(*
SPDX-FileCopyrightText: c 2026 Oleksandr Tiutyk <trofimich@gmail.com>
SPDX-License-Identifier: MIT
License: https://opensource.org/license/mit
*)

(*!
<summary>Groups fixed-capacity list copying, borrowing, editing, search, sorting and overflow cases.</summary>
<description>
Owns the cases, their fixed registration array and any fixtures borrowed by the cases.
Each borrowed fixture is reserved for its case throughout the group lifetime. Use from one task at a stable address.
</description>
*)

{attribute 'no_assign'}
{attribute 'no_explicit_call' := 'do not call this function block directly'}
FUNCTION_BLOCK StaticListTestGroup EXTENDS TOF_Testing.TestGroup<16>
VAR_STAT
	{attribute 'hide'}
	_ClassName : STRING := __POUNAME();
END_VAR
VAR
	_AppendList : TOF_Collections.List<8>(valueValidator := 0);
	_InsertList : TOF_Collections.List<8>(valueValidator := 0);
	_GetAndSetList : TOF_Collections.List<8>(valueValidator := 0);
	_FindList : TOF_Collections.List<8>(valueValidator := 0);
	_ContainsList : TOF_Collections.List<8>(valueValidator := 0);
	_ContainsGenericList : TOF_Collections.List<8>(valueValidator := 0);
	_RemoveFirstList : TOF_Collections.List<8>(valueValidator := 0);
	_RemoveMatchedList : TOF_Collections.List<8>(valueValidator := 0);
	_RemoveAtList : TOF_Collections.List<8>(valueValidator := 0);
	_SwapList : TOF_Collections.List<8>(valueValidator := 0);
	_AppendGenericList : TOF_Collections.List<8>(valueValidator := 0);
	_InsertGenericList : TOF_Collections.List<8>(valueValidator := 0);
	_GetAndSetGenericList : TOF_Collections.List<8>(valueValidator := 0);

	_Append : ListAppendTest(name := "Append", parent := THIS^, list := _AppendList);
	_Insert : ListInsertTest(name := "Insert", parent := THIS^, list := _InsertList);
	_GetAndSet : ListGetAndSetTest(name := "GetAndSet", parent := THIS^, list := _GetAndSetList);
	_Find : ListFindTest(name := "Find", parent := THIS^, list := _FindList);
	_Contains : ListContainsTest(name := "Contains", parent := THIS^, list := _ContainsList);
	_ContainsGeneric : ListContainsGenericTest(name := "ContainsGeneric", parent := THIS^, list := _ContainsGenericList);
	_RemoveFirst : ListRemoveFirstTest(name := "RemoveFirst", parent := THIS^, list := _RemoveFirstList);
	_RemoveMatched : ListRemoveMatchedTest(name := "RemoveMatched", parent := THIS^, list := _RemoveMatchedList);
	_RemoveAt : ListRemoveAtTest(name := "RemoveAt", parent := THIS^, list := _RemoveAtList);
	_Swap : ListSwapTest(name := "Swap", parent := THIS^, list := _SwapList);
	_Sort : StaticListSortTest(name := "Sort", parent := THIS^);
	_AppendGeneric : ListAppendGenericTest(name := "AppendGeneric", parent := THIS^, list := _AppendGenericList);
	_InsertGeneric : ListInsertGenericTest(name := "InsertGeneric", parent := THIS^, list := _InsertGenericList);
	_GetAndSetGeneric : ListGetAndSetGenericTest(
		name := "GetAndSetGeneric",
		parent := THIS^,
		list := _GetAndSetGenericList
	);
	_Clear : StaticListClearTest(name := "Clear", parent := THIS^);
	_Overflow : StaticListOverflowTest(name := "Overflow", parent := THIS^);

	_Children : ARRAY [0.._ChildCount - 1] OF TOF_Testing.ITestElement :=
	[
		_Append,
		_Insert,
		_GetAndSet,
		_Find,
		_Contains,
		_ContainsGeneric,
		_RemoveFirst,
		_RemoveMatched,
		_RemoveAt,
		_Swap,
		_Sort,
		_AppendGeneric,
		_InsertGeneric,
		_GetAndSetGeneric,
		_Clear,
		_Overflow
	];
END_VAR

//! <summary>Borrows the fixed child array. Callers must not modify it.</summary>
{attribute 'monitoring' := 'call'}
PROPERTY Children : REFERENCE TO ARRAY [0.._ChildCount - 1] OF TOF_Testing.ITestElement
GET
Children REF= _Children;
END_GET
END_PROPERTY

//! <summary>Borrows the concrete class name. Callers must not modify it.</summary>
{attribute 'monitoring' := 'call'}
PROPERTY ClassName : REFERENCE TO STRING
GET
ClassName REF= _ClassName;
END_GET
END_PROPERTY

//! <summary>Borrows the compiler-initialized namespace name. Callers must not modify it.</summary>
{attribute 'monitoring' := 'call'}
PROPERTY NamespaceName : REFERENCE TO STRING
GET
NamespaceName REF= CurrentNamespace.Name;
END_GET
END_PROPERTY

//! <summary>Reports the concrete instance size in bytes.</summary>
{attribute 'monitoring' := 'call'}
PROPERTY SelfSize : ULINT
GET
SelfSize := XSIZEOF(THIS^);
END_GET
END_PROPERTY

END_FUNCTION_BLOCK

(* stored: Version 1.1.0.1
   POU StaticListTestGroup: Id {5389c658-e0fc-4c89-81f8-525b97bf6c9f}, SpecialFunc None
   Property Children: Id {1fc68d15-e9f1-4bfe-9733-440331956d59}
   Get Get: Id {eab20938-bded-4a57-88ef-0f0fb0cbd6bd}
   Property ClassName: Id {87c73642-5bf6-431b-8bff-d107cebfeada}
   Get Get: Id {f3061394-8c44-40be-a295-97f756388c0a}
   Property NamespaceName: Id {24a22fe2-c2db-416b-9358-523ae6698ce7}
   Get Get: Id {1680da9d-5301-4a3c-a798-9be4fbb726d6}
   Property SelfSize: Id {d74794c6-f6e0-4858-9c71-f79af8848a04}
   Get Get: Id {ddfe4ffc-186a-4e9f-a9d8-505b8ff9ec50} *)
